(* IEC 61131-3 sources: kns-port-domestic/upstream/kns-pump-station/src/POUs/Station/FB_PowerRestore, 2 files *)

(* ---- FB_PowerRestore.decl.st ---- *)
// Назначение: питание и последовательный пуск (04 §13). Первый вызов — «задержка» tPlcStart
//             (выходы устройств ещё не посчитаны: xPowerOk первого вызова не используется);
//             напряжение пропало — «нет напряжения», запросов нет (событие 101008); вернулось —
//             «задержка» tPwrRestart (событие 101009); затем шаги: разрешён k-й запрос, следующий —
//             через tSeqStep после подтверждения k пусков или через STN_SEQ_START_TIMEOUT, если пуск
//             не подтвердился (АВР уже назначил замену); конец — разрешено не меньше требуемого
//             (событие 101010, значение — число разрешённых пусков).
// Автор:      kr0nsch
// Версия:     0.1.0
// Документ:   docs/DESIGN.md, раздел 6.9; docs/04_algorithms.md, раздел 13
FUNCTION_BLOCK FB_PowerRestore
VAR_INPUT
    xPowerOk           : BOOL;      // fbES301.xValue (подтверждение 3 с — задержка DI)
    uiRequired         : UINT;      // от действующего управления
    uiRunningRequested : UINT;      // FB_PumpRotation: запрошены и работают
    itfTime            : PL.I_TimeSource;
    itfEvents          : I_StationEventSink;
END_VAR
VAR_IN_OUT CONSTANT
    stCfg : ST_StationCfg;          // tPwrRestart, tSeqStep, tPlcStart
END_VAR
VAR_OUTPUT
    xPowerLost     : BOOL;
    xRestart       : BOOL;          // задержка после восстановления (старта) или последовательный пуск
    uiRequestLimit : UINT;          // 0 — нет запросов; k — шаг k; STN_PUMP_COUNT — без ограничения
    uiSeqRemain_s  : UINT;          // до следующего шага, с (вверх)
END_VAR
VAR
    xFirstCall   : BOOL := TRUE;    // первый вызов: задержка tPlcStart
    xLost        : BOOL;            // состояние «нет напряжения»
    xDelay       : BOOL;            // состояние «задержка» (после старта или восстановления)
    xPlcStart    : BOOL;            // задержка — после старта ПЛК (tPlcStart), иначе tPwrRestart
    xSeq         : BOOL;            // состояние «последовательный пуск»
    uiStep       : UINT;            // разрешено запросов на шаге
    xConfirmed   : BOOL;            // пуски шага подтверждены (отсчёт tSeqStep)
    fbDelay      : PL.FB_Delay;     // задержка tPlcStart / tPwrRestart
    fbStepWait   : PL.FB_Delay;     // tSeqStep после подтверждения пусков шага
    fbStepTimeout : PL.FB_Delay;    // пуск шага не подтвердился за STN_SEQ_START_TIMEOUT
END_VAR
VAR_TEMP
    xAdvance  : BOOL;               // перейти к следующему шагу
    tRemain   : TIME;               // до следующего шага
    udiRemain : UDINT;              // то же, с (вверх)
END_VAR

(* ---- FB_PowerRestore.impl.st ---- *)
// 1. Переходы по питанию (диаграмма 04 §13.2). В первом вызове xPowerOk ещё не посчитан
//    устройством (станция вызывается до PRG_Devices): старт ПЛК — сразу «задержка» tPlcStart
IF xFirstCall THEN
    xDelay := TRUE;
    xPlcStart := TRUE;
    xLost := FALSE;
    xSeq := FALSE;
    IF itfEvents <> 0 THEN
        itfEvents.LogEvent(eEvent := E_StationEvent.RestartBegin, rValue := 0.0);
    END_IF
ELSIF NOT xPowerOk THEN
    IF NOT xLost THEN
        xLost := TRUE;
        xDelay := FALSE;
        xSeq := FALSE;
        IF itfEvents <> 0 THEN
            itfEvents.LogEvent(eEvent := E_StationEvent.PowerLost, rValue := 0.0);
        END_IF
    END_IF
ELSIF xLost THEN
    xLost := FALSE;
    xDelay := TRUE;
    xPlcStart := FALSE;
    IF itfEvents <> 0 THEN
        itfEvents.LogEvent(eEvent := E_StationEvent.RestartBegin, rValue := 0.0);
    END_IF
END_IF

// 2. Задержка после старта или восстановления; затем первый шаг
fbDelay(xIn := xDelay, tOnDelay := SEL(xPlcStart, stCfg.tPwrRestart, stCfg.tPlcStart), itfTime := itfTime);
IF xDelay AND fbDelay.xOut THEN
    xDelay := FALSE;
    xSeq := TRUE;
    uiStep := 1;
    xConfirmed := FALSE;
    fbStepWait.Preset(xValue := FALSE);
    fbStepTimeout.Preset(xValue := FALSE);
END_IF

// 3. Шаги: следующий запрос — через tSeqStep после подтверждения пусков шага (ОС), либо через
//    STN_SEQ_START_TIMEOUT, если пуск не подтвердился
IF xSeq AND NOT xConfirmed AND uiRunningRequested >= uiStep THEN
    xConfirmed := TRUE;
END_IF
fbStepWait(xIn := xSeq AND xConfirmed, tOnDelay := stCfg.tSeqStep, itfTime := itfTime);
fbStepTimeout(xIn := xSeq AND NOT xConfirmed, tOnDelay := GVL_Const.STN_SEQ_START_TIMEOUT, itfTime := itfTime);
xAdvance := xSeq AND uiStep < uiRequired AND (fbStepWait.xOut OR fbStepTimeout.xOut);
IF xAdvance THEN
    uiStep := uiStep + 1;
    xConfirmed := FALSE;
    fbStepWait.Preset(xValue := FALSE);
    fbStepTimeout.Preset(xValue := FALSE);
END_IF
IF xSeq AND uiStep >= uiRequired AND (uiRunningRequested >= uiRequired OR fbStepTimeout.xOut) THEN
    // разрешено не меньше требуемого и все запрошенные пущены (или пуск шага не подтвердился за
    // STN_SEQ_START_TIMEOUT) — последовательность завершена. Только «разрешено не меньше требуемого» мало:
    // после Restart автоматика набирает потребность заново, и в конце задержки она ещё не полная (PMI-34)
    xSeq := FALSE;
    IF itfEvents <> 0 THEN
        itfEvents.LogEvent(eEvent := E_StationEvent.RestartDone, rValue := UINT_TO_REAL(MIN(uiStep, uiRequired)));
    END_IF
END_IF

// 4. Выходы
xPowerLost := xLost;
xRestart := xDelay OR xSeq;
IF xLost OR xDelay THEN
    uiRequestLimit := 0;
ELSIF xSeq THEN
    uiRequestLimit := uiStep;
ELSE
    uiRequestLimit := GVL_Const.STN_PUMP_COUNT;
END_IF

// остаток до следующего шага в целых секундах вверх (HMI, 04 §13.2)
tRemain := T#0S;
IF xDelay THEN
    tRemain := fbDelay.tRemaining;
ELSIF xSeq AND xConfirmed THEN
    tRemain := fbStepWait.tRemaining;
ELSIF xSeq THEN
    tRemain := fbStepTimeout.tRemaining;
END_IF
udiRemain := TIME_TO_UDINT(tRemain) / GVL_Const.STN_MS_PER_S;
IF udiRemain * GVL_Const.STN_MS_PER_S < TIME_TO_UDINT(tRemain) THEN
    udiRemain := udiRemain + 1;
END_IF
uiSeqRemain_s := UDINT_TO_UINT(MIN(udiRemain, UINT_TO_UDINT(PL.GVL_Const.UINT_MAX)));
xFirstCall := FALSE;
